Fanuc KAREL source: kt00518.KL

PROGRAM KT00518
%STACKSIZE=65535
%PRIORITY=65535
%NOLOCKGROUP
VAR
P1 : XYZWPREXT
P2 : XYZWPR
OUT : BOOLEAN
BEGIN
P1.X=1.0
P2.Y=2.0
-- UNRESOLVED_PC line 10 opcodes [49 7E 49 7E AC 23] marker_code=40
END KT00518
